// TIA Portal V20 export
Screen "Pop-up_Opmodes12_Popup"  645x267
  ScreenItem "Background" at 0,0 size 645x267  Type=HmiRectangle
  ScreenItem "Descr_HmiPanel" at 1,208 size 56x40  Type=HmiTextBox
  ScreenItem "Linie1_LightGrey" at 10,207 size 520x0  Type=HmiLine
  ScreenItem "Linie1_DarkGrey" at 10,207 size 520x0  Type=HmiLine
  ScreenItem "Linie1_LightGrey_1" at 10,249 size 520x0  Type=HmiLine
  ScreenItem "Linie1_DarkGrey_1" at 10,248 size 520x0  Type=HmiLine
  ScreenItem "Overview_OPMode" at 1,1 size 643x25  Type=HmiTextBox
  ScreenItem "Descr_OPMode" at 1,26 size 550x40  Type=HmiTextBox
  ScreenItem "OPMode12_small" at 540,136 size 90x60  Type=HmiButton
  ScreenItem "OPMode1_small" at 15,71 size 90x60  Type=HmiButton
  ScreenItem "OPMode2_small" at 15,136 size 90x60  Type=HmiButton
  ScreenItem "OPMode3_small" at 120,71 size 90x60  Type=HmiButton
  ScreenItem "OPMode5_small" at 225,71 size 90x60  Type=HmiButton
  ScreenItem "OPMode4_small" at 121,136 size 90x60  Type=HmiButton
  ScreenItem "OPMode6_small" at 226,136 size 90x60  Type=HmiButton
  ScreenItem "OPMode7_small" at 330,71 size 90x60  Type=HmiButton
  ScreenItem "OPMode8_small" at 331,136 size 90x60  Type=HmiButton
  ScreenItem "OPMode9_small" at 435,71 size 90x60  Type=HmiButton
  ScreenItem "OPMode10_small" at 435,136 size 90x60  Type=HmiButton
  ScreenItem "OPMode11_small" at 540,71 size 90x60  Type=HmiButton
  ScreenItem "OPMode1_wide" at 10,71 size 100x60  Type=HmiButton
  ScreenItem "OPMode2_wide" at 10,136 size 100x60  Type=HmiButton
  ScreenItem "OPMode3_wide" at 115,71 size 100x60  Type=HmiButton
  ScreenItem "OPMode4_wide" at 116,136 size 100x60  Type=HmiButton
  ScreenItem "OPMode5_wide" at 220,71 size 100x60  Type=HmiButton
  ScreenItem "OPMode6_wide" at 221,136 size 100x60  Type=HmiButton
  ScreenItem "OPMode7_wide" at 326,71 size 100x60  Type=HmiButton
  ScreenItem "OPMode8_wide" at 326,136 size 100x60  Type=HmiButton
  ScreenItem "OPMode9_wide" at 430,71 size 100x60  Type=HmiButton
  ScreenItem "OPMode10_wide" at 430,136 size 100x60  Type=HmiButton
  ScreenItem "OPMode11_wide" at 535,71 size 100x60  Type=HmiButton
  ScreenItem "OPMode12_wide" at 535,136 size 100x60  Type=HmiButton
  ScreenItem "Overview_HMI-OP" at 554,207 size 90x60  Type=HmiButton
  ScreenItem "Cancel Mode" at 554,1 size 90x60  Type=HmiButton
  ScreenItem "OPMode1_Foreground_Blocked" at 10,71 size 100x60  Type=HmiGraphicView
  ScreenItem "OPMode2_Foreground_Blocked" at 10,136 size 100x60  Type=HmiGraphicView
  ScreenItem "OPMode3_Foreground_Blocked" at 115,71 size 100x60  Type=HmiGraphicView
  ScreenItem "OPMode4_Foreground_Blocked" at 115,136 size 100x60  Type=HmiGraphicView
  ScreenItem "OPMode5_Foreground_Blocked" at 220,71 size 100x60  Type=HmiGraphicView
  ScreenItem "OPMode6_Foreground_Blocked" at 221,136 size 100x60  Type=HmiGraphicView
  ScreenItem "OPMode7_Foreground_Blocked" at 326,71 size 100x60  Type=HmiGraphicView
  ScreenItem "OPMode8_Foreground_Blocked" at 326,136 size 100x60  Type=HmiGraphicView
  ScreenItem "OPMode9_Foreground_Blocked" at 430,71 size 100x60  Type=HmiGraphicView
  ScreenItem "OPMode10_Foreground_Blocked" at 430,136 size 100x60  Type=HmiGraphicView
  ScreenItem "OPMode11_Foreground_Blocked" at 535,71 size 100x60  Type=HmiGraphicView
  ScreenItem "OPMode12_Foreground_Blocked" at 535,136 size 100x60  Type=HmiGraphicView
  ScreenItem "OPMode1_Blocked" at 93,75 size 14x14  Type=HmiGraphicView
  ScreenItem "OPMode2_Blocked" at 93,139 size 14x14  Type=HmiGraphicView
  ScreenItem "OPMode3_Blocked" at 199,75 size 14x14  Type=HmiGraphicView
  ScreenItem "OPMode4_Blocked" at 199,139 size 14x14  Type=HmiGraphicView
  ScreenItem "OPMode5_Blocked" at 303,75 size 14x14  Type=HmiGraphicView
  ScreenItem "OPMode6_Blocked" at 305,139 size 14x14  Type=HmiGraphicView
  ScreenItem "OPMode7_Blocked" at 408,75 size 14x14  Type=HmiGraphicView
  ScreenItem "OPMode8_Blocked" at 408,139 size 14x14  Type=HmiGraphicView
  ScreenItem "OPMode9_Blocked" at 514,75 size 14x14  Type=HmiGraphicView
  ScreenItem "OPMode10_Blocked" at 514,139 size 14x14  Type=HmiGraphicView
  ScreenItem "OPMode11_Blocked" at 618,75 size 14x14  Type=HmiGraphicView
  ScreenItem "OPMode12_Blocked" at 618,139 size 14x14  Type=HmiGraphicView
